Staubli VAL3: main.pgx

public program main()
  local bool l_bExit
  local bool l_bResult
  local num l_nTool
  local tool l_tTool
  local num l_nUsingLib
  local num l_nResult
  local string l_sLib
  local num i
begin
  do
    if util:sPage!="setting"
      util:sPage="setting"
      call util:loadingPage()
      call onStart()
      call bind()
      userPage("setting")
      delay(0.5)
    endIf

    if sSelTool != sLastTool
      sLastTool=sSelTool
      toNum(sLastTool,l_nTool,l_bResult)
    endIf
    if bTeach
      bTeach=false
      call teachHome()
    elseIf bMove
      bMove=false
      call moveTohome()
    elseIf bSetup
      bSetup=false
      if l_nTool!=savedata:nJogTool
        savedata:nJogTool=l_nTool
        call savedata:setBaseJOG(l_nTool)
        savedata:libSave()
        delay(0.1)
      endIf
    elseIf bChangeLib
      bChangeLib=false
      if workingMode()!=1
        popUpMsg("请先将工作模式切换到手动模式")
      else
        l_sLib=delete(sUsingLib,3,0)
        toNum(l_sLib,l_nUsingLib,l_bResult)
        if !l_bResult
          return
        else
          bIsDoing=true
          savedata:nLibIndex=l_nUsingLib
          savedata:libSave()

          bToSave=true
          call prog:onSave(bToSave)
          bToSave=true
          call trajectory:onSave(bToSave)
          logMsg("手动开始切换:"+toString(".2",clock()))
          call prog:loadPROG(l_nUsingLib,l_nResult)
          call trajectory:loadTRAJ(l_nUsingLib,l_nResult)

          bIsDoing=false
        endIf
      endIf
    elseIf bBack
      bBack=false
      l_bExit=true
    endIf

    call libTqe:refresh()
    //    if bLock==true
    //      sBtnUnLock="解锁"
    //    else
    //      sBtnUnLock="保存"
    //    endIf
    delay(0)
  until l_bExit==true
end
